(* IEC 61131-3 sources: building-irrigation-scada/PLC/Codesys/Zone03, 2 files *)

(* ---- FB_IrrigationZone.declaration.reference.st ---- *)
(*
Source reference: Zone03 / CODESYS / FB_IrrigationZone declaration
Recovered from: docs/plc-source-reference-baseline
Verification: NOT VERIFIED against the current native CODESYS application
Native project: intentionally not included in this repository
*)
FUNCTION_BLOCK FB_IrrigationZone
VAR_INPUT
    xCmdStart           : BOOL;   (* momentary/latched command from SCADA, cleared after use *)
    xCmdStop             : BOOL;
    xCmdFaultReset       : BOOL;
    xAuto                : BOOL;  (* TRUE = automatic moisture-threshold control *)
    xSimEnable           : BOOL;  (* master enable — nothing runs while FALSE *)
    xSimCommFault        : BOOL;
    xSimActuatorFault    : BOOL;
    xSimSensorFault      : BOOL;
    xSimRestriction      : BOOL;
    rMoistureLowSP       : REAL;
    rMoistureHighSP      : REAL;
    rSimFlowTarget       : REAL;
    rSimFlowRate         : REAL;
    rSimMoistureRate     : REAL;
    rSimDryRate          : REAL;
    rSimLowFlowLimit     : REAL;
END_VAR
VAR_OUTPUT
    xRunning             : BOOL;
    xRunFeedback         : BOOL;
    xFault                : BOOL;
    xPermissive          : BOOL;
    xFlowOK              : BOOL;
    xProcessOK           : BOOL;
    xCommanded           : BOOL;
    xAutoActive          : BOOL;
    xManual              : BOOL;
    xLowFlow             : BOOL;
    xCommOK              : BOOL;
    xSimActive           : BOOL;
    rFlow                : REAL;
    rMoisture            : REAL;
    rValvePosition       : REAL;  (* 0.0-100.0 *)
    udiTotalRuntimeSec   : UDINT;
END_VAR
VAR
    xFaultLatch          : BOOL;
    xAutoDemand          : BOOL;
    rFlowTarget          : REAL;
    rFlowError           : REAL;
    rFlowStep            : REAL;
    rMoistureStep        : REAL;
    uiRuntimeTicks       : UINT;
    rtStart              : R_TRIG;
    rtStop               : R_TRIG;
    rtFaultReset         : R_TRIG;
    fbTick               : TON;
END_VAR

(* ---- FB_IrrigationZone.implementation.reference.st ---- *)
(*
Source reference: Zone03 / CODESYS / FB_IrrigationZone implementation
Recovered from: docs/plc-source-reference-baseline
Verification: NOT VERIFIED against the current native CODESYS application
Native project: intentionally not included in this repository
The implementation body below is retained without logic changes.
*)

// =============================================================
// 1. COMMAND EDGE DETECTION
// =============================================================
rtStart(CLK := xCmdStart);
rtStop(CLK := xCmdStop);
rtFaultReset(CLK := xCmdFaultReset);

// =============================================================
// 2. STATUS MIRRORS
// =============================================================
xSimActive := xSimEnable;
xCommOK    := NOT xSimCommFault;

// =============================================================
// 3. FAULT GENERATION / RESET
// =============================================================
IF xSimActuatorFault OR xSimSensorFault THEN
    xFaultLatch := TRUE;
END_IF;

IF rtFaultReset.Q THEN
    IF NOT xSimActuatorFault AND NOT xSimSensorFault THEN
        xFaultLatch := FALSE;
    END_IF;
END_IF;

// =============================================================
// 4. PERMISSIVE
//    NOTE: requires xSimEnable = TRUE. If nothing is running and
//    everything else looks correctly wired, check this input first.
// =============================================================
xPermissive :=
    NOT xFaultLatch
    AND NOT xSimActuatorFault
    AND NOT xSimSensorFault
    AND xCommOK
    AND xSimEnable;

// =============================================================
// 5. AUTO DEMAND (hysteresis on moisture, does not touch xRunning directly)
// =============================================================
IF rMoisture <= rMoistureLowSP THEN
    xAutoDemand := TRUE;
ELSIF rMoisture >= rMoistureHighSP THEN
    xAutoDemand := FALSE;
END_IF;
// else: holds previous state — this is the intended dead-band behavior

// =============================================================
// 6. RUNNING DECISION
//    Fix: Stop always wins, even in Auto mode, for the scan it's pressed.
// =============================================================
xAutoActive := FALSE;

IF xAuto AND xPermissive THEN
    xAutoActive := TRUE;
    xRunning    := xAutoDemand;
ELSIF xPermissive THEN
    IF rtStart.Q THEN
        xRunning := TRUE;
    END_IF;
END_IF;

// Manual/safety Stop — always evaluated last, always wins this scan,
// regardless of Auto/Manual mode.
IF rtStop.Q THEN
    xRunning    := FALSE;
    xAutoDemand := FALSE;
END_IF;

// =============================================================
// 7. FAULT / COMMUNICATION / ENABLE SAFETY
// =============================================================
IF xFaultLatch THEN
    xRunning := FALSE;
END_IF;

IF NOT xCommOK THEN
    xRunning := FALSE;
END_IF;

IF NOT xSimEnable THEN
    xRunning := FALSE;
END_IF;

// =============================================================
// 8. PROCESS COMMAND
// =============================================================
xCommanded := xRunning AND xPermissive;

// =============================================================
// 9. 100 ms SIMULATION TICK
// =============================================================
fbTick(IN := TRUE, PT := T#100MS);

IF fbTick.Q THEN
    fbTick(IN := FALSE);   // retrigger for next 100 ms interval

    // ---- Valve ----
    IF xCommanded THEN
        rValvePosition := 100.0;
    ELSE
        rValvePosition := 0.0;
    END_IF;

    // ---- Flow target ----
    IF xCommanded THEN
        rFlowTarget := rSimFlowTarget;
        IF xSimRestriction THEN
            rFlowTarget := rFlowTarget * 0.25;
        END_IF;
    ELSE
        rFlowTarget := 0.0;
    END_IF;

    // ---- Flow ramp ----
    rFlowError := rFlowTarget - rFlow;
    rFlowStep  := ABS(rSimFlowRate) * 0.1;
    IF rFlowStep < 0.1 THEN
        rFlowStep := 0.1;
    END_IF;

    IF rFlowError > rFlowStep THEN
        rFlow := rFlow + rFlowStep;
    ELSIF rFlowError < -rFlowStep THEN
        rFlow := rFlow - rFlowStep;
    ELSE
        rFlow := rFlowTarget;
    END_IF;

    IF rFlow < 0.0 THEN
        rFlow := 0.0;
    END_IF;

    IF xSimSensorFault THEN
        rFlow := 0.0;   // sensor fault -> invalid/zero feedback
    END_IF;

    // ---- Moisture process ----
    IF xCommanded AND (rFlow > 0.0) THEN
        rMoistureStep := ABS(rSimMoistureRate) * 0.1;
        rMoisture     := rMoisture + rMoistureStep;
    ELSE
        rMoistureStep := ABS(rSimDryRate) * 0.1;
        rMoisture     := rMoisture - rMoistureStep;
    END_IF;

    IF rMoisture > 100.0 THEN rMoisture := 100.0; END_IF;
    IF rMoisture < 0.0   THEN rMoisture := 0.0;   END_IF;

    // ---- Flow quality ----
    xFlowOK := TRUE;
    IF xCommanded AND (rFlow < rSimLowFlowLimit) THEN
        xFlowOK := FALSE;
    END_IF;

    xLowFlow    := xCommanded AND NOT xFlowOK;
    xProcessOK  := xPermissive AND xFlowOK;

    // ---- Runtime accumulation ----
    IF xRunning THEN
        uiRuntimeTicks := uiRuntimeTicks + 1;
        IF uiRuntimeTicks >= 10 THEN   // 10 x 100ms = 1s
            udiTotalRuntimeSec := udiTotalRuntimeSec + 1;
            uiRuntimeTicks := 0;
        END_IF;
    END_IF;
END_IF;

// =============================================================
// 10. OUTPUT MAPPING
// =============================================================
xRunFeedback := xRunning;
xFault       := xFaultLatch;
xManual      := NOT xAuto;

// =============================================================
// 11. COMMAND CONSUMPTION
//     Momentary PLC-side commands are cleared by the CALLING program
//     (the GVL write-back happens where this FB is instantiated —
//     see the wiring example below), not inside the FB itself, so the
//     FB stays reusable and doesn't reach into a specific GVL.
// =============================================================
